// Commande de déploiement (docs/05 § 10)
{attribute 'qualified_only'}
{attribute 'strict'}
TYPE E_DeployCmd :
(
    None := 0,
    Verify := 1,
    Activate := 2,
    Cancel := 3
) USINT;
END_TYPE

(* stored: Version 1.1.0.1, ProductVersion 3.1.4024.12
   DUT E_DeployCmd: Id {966a08f5-4c28-505f-ae95-e6a3a32f2fba} *)
